// TIA Portal V21 export
// export: Created 2026-08-21T20:18:53.5971282Z, ExportSetting None, DisplayName Totally Integrated Automation Portal, DisplayVersion V21, DisplayName STEP 7 Professional, DisplayVersion V21, DisplayName STEP 7 Safety, DisplayVersion V21, DisplayName Tech WebApplication, DisplayVersion V21, DisplayName WinCC Basic/Comfort/Advanced, DisplayVersion V21, DisplayName WinCC Professional, DisplayVersion V21, DisplayName WinCC Unified, DisplayVersion V21
FUNCTION "BoolToDigVal_1" : Void   // FC19, SCL
{ S7_Optimized_Access := 'TRUE' }
// stored: SetENOAutomatically false
   VAR_INPUT
      In : Bool;
      ST : Byte;
   END_VAR
   VAR_OUTPUT
      Out : "DigVal";
   END_VAR
BEGIN
   #Out.ST := #ST;
   #Out.Value := #In;
END_FUNCTION
